FUNCTION_BLOCK RP (* Basic Function Block Type *)
  (* Standard: 61499-2 *)
  (* Version 0.0, 1/4/2020, prana, nxtControl GmbH, Template *)
  PACKAGE Main;
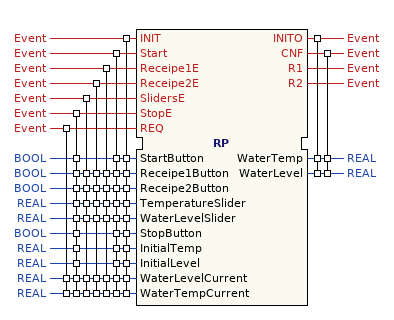
  EVENT_INPUT
    INIT WITH StartButton, Receipe1Button, Receipe2Button, TemperatureSlider, WaterLevelSlider, StopButton, InitialTemp, InitialLevel, WaterLevelCurrent, WaterTempCurrent;
    Start WITH StartButton, Receipe1Button, Receipe2Button, TemperatureSlider, WaterLevelSlider, StopButton, InitialTemp, InitialLevel, WaterLevelCurrent, WaterTempCurrent;
    Receipe1E WITH Receipe1Button, Receipe2Button, TemperatureSlider, WaterLevelSlider, WaterLevelCurrent, WaterTempCurrent; (* Initialization Request *)
    Receipe2E WITH Receipe1Button, Receipe2Button, TemperatureSlider, WaterLevelSlider, WaterLevelCurrent, WaterTempCurrent; (* Normal Execution Request *)
    SlidersE WITH Receipe1Button, Receipe2Button, TemperatureSlider, WaterLevelSlider, WaterLevelCurrent, WaterTempCurrent;
    StopE WITH StartButton, Receipe1Button, Receipe2Button, TemperatureSlider, WaterLevelSlider, StopButton, InitialTemp, InitialLevel, WaterLevelCurrent, WaterTempCurrent;
    REQ WITH WaterLevelCurrent, WaterTempCurrent;
  END_EVENT
  EVENT_OUTPUT
    INITO WITH WaterLevel, WaterTemp; (* Initialization Confirm *)
    CNF WITH WaterLevel, WaterTemp; (* Execution Confirmation *)
    R1;
    R2;
  END_EVENT
  VAR_INPUT
    StartButton : BOOL;
    Receipe1Button : BOOL; (* Input event qualifier *)
    Receipe2Button : BOOL;
    TemperatureSlider : REAL;
    WaterLevelSlider : REAL;
    StopButton : BOOL;
    InitialTemp : REAL;
    InitialLevel : REAL;
    WaterLevelCurrent : REAL;
    WaterTempCurrent : REAL;
  END_VAR
  VAR_OUTPUT
    WaterTemp : REAL;
    WaterLevel : REAL; (* Output event qualifier *)
  END_VAR
  VAR
    X1 : REAL := 165.50;
    Y1 : REAL := 50.00;
    X2 : REAL := 250.50;
    Y2 : REAL := 68.96;
  END_VAR
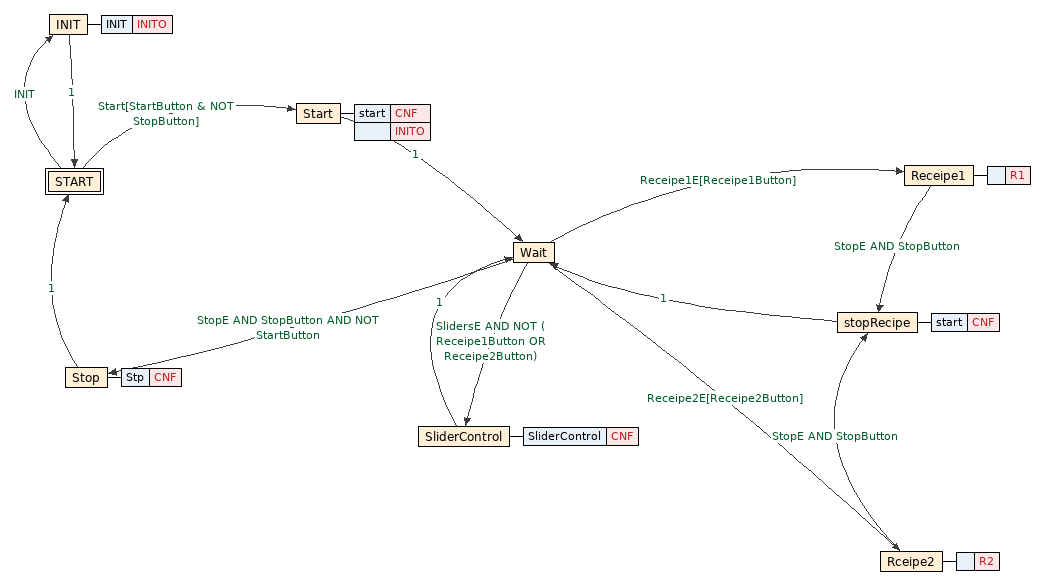
  EC_STATES
    START; (* Initial State *)
    SliderControl : SliderControl -> CNF;
    Start : start -> CNF, -> INITO;
    Wait;
    Stop : Stp -> CNF;
    INIT : INIT -> INITO;
    Receipe1 : -> R1;
    Rceipe2 : -> R2;
    stopRecipe : start -> CNF;
  END_STATES
  EC_TRANSITIONS
    Wait TO SliderControl := SlidersE AND NOT ( Receipe1Button OR Receipe2Button);
    SliderControl TO Wait := 1;
    START TO Start := Start[StartButton & NOT StopButton];
    Start TO Wait := 1;
    Wait TO Stop := StopE AND StopButton AND NOT StartButton;
    Stop TO START := 1;
    START TO INIT := INIT;
    INIT TO START := 1;
    Wait TO Receipe1 := Receipe1E[Receipe1Button];
    Wait TO Rceipe2 := Receipe2E[Receipe2Button];
    Receipe1 TO stopRecipe := StopE AND StopButton;
    Rceipe2 TO stopRecipe := StopE AND StopButton;
    stopRecipe TO Wait := 1;
  END_TRANSITIONS
  ALGORITHM INIT IN ST: (* Initialization algorithm *)
;
  END_ALGORITHM
  ALGORITHM SliderControl IN ST:
WaterLevel := WaterLevelSlider;
WaterTemp := TemperatureSlider;
  END_ALGORITHM
  ALGORITHM start IN ST:
WaterLevel := InitialLevel;
WaterTemp := InitialTemp;
  END_ALGORITHM
  ALGORITHM Stp IN ST:
WaterLevel := 0;
WaterTemp := 0;
  END_ALGORITHM
  ALGORITHM X1 IN ST:
WaterLevel := X1;
WaterTemp := Y2;
  END_ALGORITHM
  ALGORITHM X2 IN ST:
WaterLevel := X2;
WaterTemp := Y2;
  END_ALGORITHM
  ALGORITHM Drain IN ST:
WaterLevel := 0;
WaterTemp := 0;
  END_ALGORITHM
END_FUNCTION_BLOCK
